(* PLC project Zwei Steuerungen, CODESYS CODESYS V3.5 SP21, author synthetisch *)
(* stored: creationDateTime 2026-10-31T10:00:00.0000000, version 1.0.0.0, modificationDateTime 2026-10-31T09:59:00.0000000, organization Comquent GmbH *)

CONFIGURATION Verpackung
  RESOURCE Application ON PLC
  END_RESOURCE
  RESOURCE Diagnose ON PLC
  END_RESOURCE
END_CONFIGURATION

CONFIGURATION Feldbus_Koppler
END_CONFIGURATION

CONFIGURATION Achspool
END_CONFIGURATION

CONFIGURATION Handling
  RESOURCE Application ON PLC
  END_RESOURCE
END_CONFIGURATION
